RESOURCE RES0 : EMB_RES_ECO
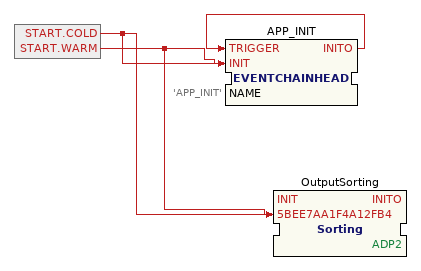
  FBS
    OutputSorting : Sorting;
    APP_INIT : EVENTCHAINHEAD(NAME := 'APP_INIT');
  END_FBS
  EVENT_CONNECTIONS
    APP_INIT.INITO TO APP_INIT.TRIGGER;
    START.COLD TO APP_INIT.INIT;
    START.WARM TO APP_INIT.INIT;
    START.COLD TO OutputSorting.5BEE7AA1F4A12FB4;
    START.WARM TO OutputSorting.5BEE7AA1F4A12FB4;
  END_CONNECTIONS
END_RESOURCE
